// TIA Portal V21 export
FUNCTION "FC_LadContacts" : Void   // FC6, LAD
TITLE = KOP-Kontakte und -Spulen / LAD contacts and coils
{ S7_Optimized_Access := 'TRUE' }
// stored: SetENOAutomatically false
   VAR_INPUT
      Start : Bool;   // Startbefehl / Start command
      Stop : Bool;   // Stoppbefehl / Stop command
      Sensor : Bool;   // Produktsensor / Product sensor
      Enable : Bool;   // Freigabe / Enable
      Reset : Bool;   // Rücksetzbefehl / Reset command
   END_VAR
   VAR_OUTPUT
      Motor : Bool;   // Motor ein / Motor on
      Pulse : Bool;   // Impuls bei steigender Flanke des Sensors / Pulse on rising edge of the sensor
      FallingPulse : Bool;   // Impuls bei fallender Flanke des Sensors / Pulse on falling edge of the sensor
      Alarm : Bool;   // Alarm wenn nicht freigegeben / Alarm when not enabled
      Lamp : Bool;   // Leuchte bei steigender Flanke der Freigabe / Lamp set on rising edge of the enable
      BranchResult : Bool;   // Ergebnis der verschachtelten Verzweigung / Result of the nested branch
   END_VAR
   VAR_IN_OUT
      Latched : Bool;   // Gespeicherter Zustand / Latched state
      RiseMemory : Bool;   // Flankenmerker steigend / Edge memory, rising
      FallMemory : Bool;   // Flankenmerker fallend / Edge memory, falling
      CoilMemory : Bool;   // Flankenmerker der Spule / Edge memory of the coil
   END_VAR
   VAR_TEMP   // added for the SCL form of the ladder/FBD networks
      _w1 : Bool;
   END_VAR
BEGIN

REGION Network 1: Schließer und Öffner / Normally open and normally closed contact
   // Der Motor läuft, solange Start gedrückt und Stopp nicht gedrückt ist. / The motor runs while start is pressed and stop is not pressed.
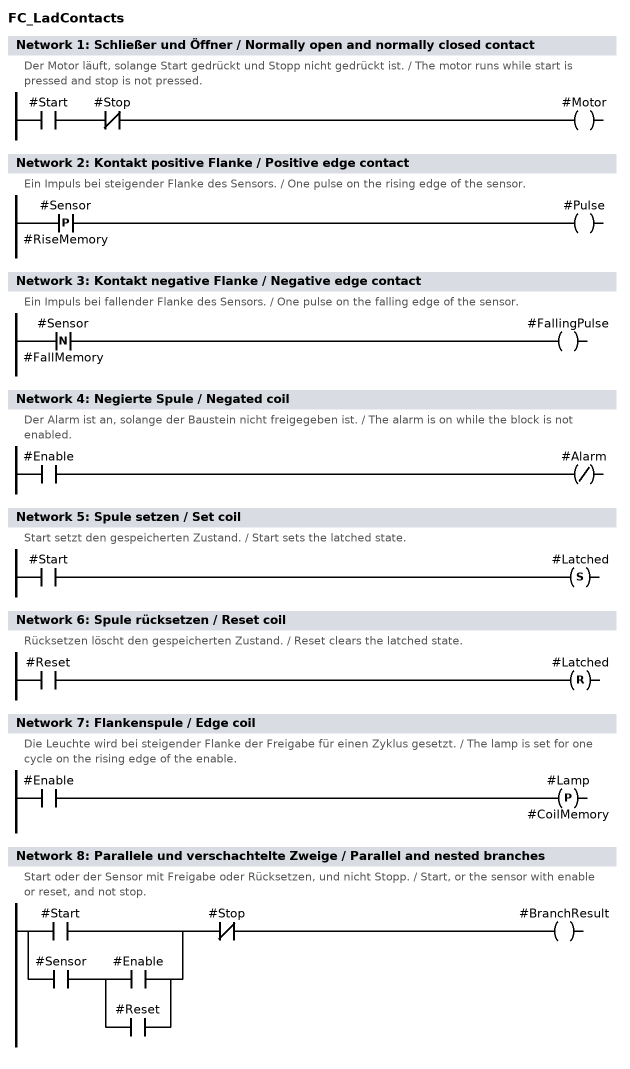
   RUNG wire#powerrail
      Contact( #Start )
      I_Contact( #Stop )
      Coil( #Motor )
   END_RUNG
   // the same network as SCL:
   #Motor := #Start AND NOT #Stop;
END_REGION

REGION Network 2: Kontakt positive Flanke / Positive edge contact
   // Ein Impuls bei steigender Flanke des Sensors. / One pulse on the rising edge of the sensor.
   RUNG wire#powerrail
      P_Contact(operand := #Sensor, bit := #RiseMemory)
      Coil( #Pulse )
   END_RUNG
   // the same network as SCL:
   #_w1 := #Sensor AND NOT #RiseMemory;   // rising edge of #Sensor
   #RiseMemory := #Sensor;
   #Pulse := #_w1;
END_REGION

REGION Network 3: Kontakt negative Flanke / Negative edge contact
   // Ein Impuls bei fallender Flanke des Sensors. / One pulse on the falling edge of the sensor.
   RUNG wire#powerrail
      N_Contact(operand := #Sensor, bit := #FallMemory)
      Coil( #FallingPulse )
   END_RUNG
   // the same network as SCL:
   #_w1 := NOT #Sensor AND #FallMemory;   // falling edge of #Sensor
   #FallMemory := #Sensor;
   #FallingPulse := #_w1;
END_REGION

REGION Network 4: Negierte Spule / Negated coil
   // Der Alarm ist an, solange der Baustein nicht freigegeben ist. / The alarm is on while the block is not enabled.
   RUNG wire#powerrail
      Contact( #Enable )
      I_Coil( #Alarm )
   END_RUNG
   // the same network as SCL:
   #Alarm := NOT #Enable;
END_REGION

REGION Network 5: Spule setzen / Set coil
   // Start setzt den gespeicherten Zustand. / Start sets the latched state.
   RUNG wire#powerrail
      Contact( #Start )
      S_Coil( #Latched )
   END_RUNG
   // the same network as SCL:
   IF #Start THEN #Latched := TRUE; END_IF;
END_REGION

REGION Network 6: Spule rücksetzen / Reset coil
   // Rücksetzen löscht den gespeicherten Zustand. / Reset clears the latched state.
   RUNG wire#powerrail
      Contact( #Reset )
      R_Coil( #Latched )
   END_RUNG
   // the same network as SCL:
   IF #Reset THEN #Latched := FALSE; END_IF;
END_REGION

REGION Network 7: Flankenspule / Edge coil
   // Die Leuchte wird bei steigender Flanke der Freigabe für einen Zyklus gesetzt. / The lamp is set for one cycle on the rising edge of the enable.
   #Lamp := #Enable AND NOT #CoilMemory;   // rising edge
   #CoilMemory := #Enable;
END_REGION

REGION Network 8: Parallele und verschachtelte Zweige / Parallel and nested branches
   // Start oder der Sensor mit Freigabe oder Rücksetzen, und nicht Stopp. / Start, or the sensor with enable or reset, and not stop.
   RUNG wire#powerrail
      Contact( #Start )
      wire#w1
      I_Contact( #Stop )
      Coil( #BranchResult )
   END_RUNG
   RUNG wire#powerrail
      Contact( #Sensor )
      wire#w2
      Contact( #Enable )
   END_RUNG wire#w1
   RUNG wire#w2
      Contact( #Reset )
   END_RUNG wire#w1
   // the same network as SCL:
   #BranchResult := (#Start OR (#Sensor AND (#Enable OR #Reset))) AND NOT #Stop;
END_REGION
END_FUNCTION
